(* Tests simple and batch log processors. *)
FUNCTION_BLOCK FB_TestLogProcessors EXTENDS FB_TestSuite

THIS^.testSimpleProcessorExportsEachRecord();
THIS^.testBatchProcessorQueuesAndFlushes();
THIS^.testProcessorsSkipBusyExporter();

(*
	The batch processor queues emitted records in arrival order (oldest at
	the head), dropping the oldest when the queue is full. Flushing moves
	the oldest maxExportBatchSize records into the exporter's queue, on a
	full batch or when the schedule delay elapses, so records leave in order
	and memory stays bounded however fast the PLC logs. queuedCount reports
	the records waiting for export, and droppedCount the records lost.

	FB_LoggerProvider.tick() unstages every processor, so a processor must be
	staged again before each tick.
*)
METHOD testBatchProcessorQueuesAndFlushes : REFERENCE TO FB_Test
VAR
	resourceA: FB_Resource('resource.a');
	resourceB: FB_Resource('resource.b');
	providerA: FB_LoggerProvider(resourceA);
	providerB: FB_LoggerProvider(resourceB);
	scopeA: FB_InstrumentationScope('scope.a', '1.0.0', '');
	scopeB: FB_InstrumentationScope('scope.b', '1.0.0', '');
	loggerAA: FB_Logger(scopeA, providerA);
	loggerAB: FB_Logger(scopeB, providerA);
	loggerBA: FB_Logger(scopeA, providerB);
	exporter: FB_LogRecordExporter_ForInspection;
	processor: FB_LogRecordProcessor_ForBatchInspection(
		maxQueueSize:=10,
		scheduledDelayMillis:=1000,
		maxExportBatchSize:=6,
		exporter:=exporter
	);
	// no exporter, so onEmit only enriches and never queues
	orphanProcessor: FB_LogRecordProcessor_ForBatchInspection(
		maxQueueSize:=10,
		scheduledDelayMillis:=1000,
		maxExportBatchSize:=6,
		exporter:=0
	);
	boundedExporter: FB_LogRecordExporter_ForInspection;
	boundedProcessor: FB_LogRecordProcessor_ForBatchInspection(
		maxQueueSize:=2,
		scheduledDelayMillis:=1000,
		maxExportBatchSize:=3,
		exporter:=boundedExporter
	);
	timerExporter: FB_LogRecordExporter_ForInspection;
	timerProcessor: FB_LogRecordProcessor_ForBatchInspection(
		maxQueueSize:=0,
		scheduledDelayMillis:=0,
		maxExportBatchSize:=3,
		exporter:=timerExporter
	);
	ts1: ULINT := 1;
	ts2: ULINT := 2;
	ts3: ULINT := 3;
	ts4: ULINT := 4;
	ts5: ULINT := 5;
	ts6: ULINT := 6;
	ts7: ULINT := 7;
	ts8: ULINT := 8;
	ts9: ULINT := 9;
	ts10: ULINT := 10;
	ts11: ULINT := 11;
	ts12: ULINT := 12;
	pRec: POINTER TO FB_LogRecord;
END_VAR
TcUnit.TEST('testBatchProcessorQueuesAndFlushes');
	// processor uses maxExportBatchSize 6 so the count-based flush trigger fires without waiting on the timer

	// --- Scenario: records queue in arrival order ---
	// emit interleaved across (resource, scope) pairs
	loggerBA.startLogRecord(severityNumber:=E_SeverityNumber.INFO).setTimestamp(ts1).emit();
	loggerAB.startLogRecord(severityNumber:=E_SeverityNumber.INFO).setTimestamp(ts2).emit();
	loggerAA.startLogRecord(severityNumber:=E_SeverityNumber.INFO).setTimestamp(ts3).emit();
	loggerBA.startLogRecord(severityNumber:=E_SeverityNumber.INFO).setTimestamp(ts4).emit();
	loggerAA.startLogRecord(severityNumber:=E_SeverityNumber.INFO).setTimestamp(ts5).emit();
	// note, it's bad practice to associate processors with multiple providers
	providerA
		.stageProcessor(processor)
		.tick();
	providerB
		.stageProcessor(processor)
		.tick();
	THIS^.AssertTrue(processor.lastOperationSucceeded, 'Expected the last emit to succeed');
	THIS^.AssertEquals_UDINT(5, processor.records.count, 'Expected five queued records');
	THIS^.AssertEquals_UDINT(5, processor.queuedCount, 'Expected queuedCount to report the five queued records');
	THIS^.AssertEquals_UDINT(0, processor.droppedCount, 'Expected droppedCount to be zero before the queue fills');

	// the queue keeps arrival order per provider, oldest at the head
	processor.records.reset();
	pRec := processor.records.next();
	THIS^.AssertTrue(pRec <> 0 AND_THEN pRec^.timestamp = 2, 'Expected queued record 1 to be ts2');
	pRec := processor.records.next();
	THIS^.AssertTrue(pRec <> 0 AND_THEN pRec^.timestamp = 3, 'Expected queued record 2 to be ts3');
	pRec := processor.records.next();
	THIS^.AssertTrue(pRec <> 0 AND_THEN pRec^.timestamp = 5, 'Expected queued record 3 to be ts5');
	pRec := processor.records.next();
	THIS^.AssertTrue(pRec <> 0 AND_THEN pRec^.timestamp = 1, 'Expected queued record 4 to be ts1');
	pRec := processor.records.next();
	THIS^.AssertTrue(pRec <> 0 AND_THEN pRec^.timestamp = 4, 'Expected queued record 5 to be ts4');
	THIS^.AssertTrue(processor.records.next() = 0, 'Expected queue iteration to be exhausted');

	// --- Scenario: a full batch flushes to the exporter in order ---
	// emit one more to reach maxExportBatchSize, triggering a flush
	loggerAB.startLogRecord(severityNumber:=E_SeverityNumber.INFO).setTimestamp(ts6).emit();
	providerA
		.stageProcessor(processor)
		.tick();
	THIS^.AssertEquals_UDINT(0, processor.records.count, 'Expected zero records left after a full batch flush');
	THIS^.AssertEquals_UDINT(0, processor.queuedCount, 'Expected queuedCount to drop to zero once the batch leaves');
	THIS^.AssertEquals_UDINT(6, exporter.records.count, 'Expected six records in the exported batch');

	// exported batch preserves arrival order
	exporter.records.reset();
	pRec := exporter.records.next();
	THIS^.AssertTrue(pRec <> 0 AND_THEN pRec^.timestamp = 2, 'Expected batch record 0 to be ts2');
	pRec := exporter.records.next();
	THIS^.AssertTrue(pRec <> 0 AND_THEN pRec^.timestamp = 3, 'Expected batch record 1 to be ts3');
	pRec := exporter.records.next();
	THIS^.AssertTrue(pRec <> 0 AND_THEN pRec^.timestamp = 5, 'Expected batch record 2 to be ts5');
	pRec := exporter.records.next();
	THIS^.AssertTrue(pRec <> 0 AND_THEN pRec^.timestamp = 1, 'Expected batch record 3 to be ts1');
	pRec := exporter.records.next();
	THIS^.AssertTrue(pRec <> 0 AND_THEN pRec^.timestamp = 4, 'Expected batch record 4 to be ts4');
	pRec := exporter.records.next();
	THIS^.AssertTrue(pRec <> 0 AND_THEN pRec^.timestamp = 6, 'Expected batch record 5 to be ts6');
	THIS^.AssertTrue(exporter.records.next() = 0, 'Expected batch iteration to be exhausted');

	// --- Scenario: a busy exporter holds records in the queue ---
	// the processor still queues records, but no batch leaves
	exporter.busy := TRUE;
	loggerAB.startLogRecord(severityNumber:=E_SeverityNumber.INFO).setTimestamp(ts7).emit();
	providerA
		.stageProcessor(processor)
		.tick();
	THIS^.AssertEquals_UDINT(1, processor.records.count, 'Expected one queued record while the exporter is busy');
	THIS^.AssertEquals_UDINT(6, exporter.records.count, 'Expected the busy exporter to keep the previous batch');

	// --- Scenario: a partial batch waits for the schedule delay ---
	// once free again, the single queued record stays until scheduledDelayMillis (1000 ms) elapses
	exporter.busy := FALSE;
	providerA
		.stageProcessor(processor)
		.tick();
	THIS^.AssertEquals_UDINT(1, processor.records.count, 'Expected the partial batch to wait for the schedule delay');
	THIS^.AssertEquals_UDINT(6, exporter.records.count, 'Expected no new batch before the schedule delay elapses');

	// --- Scenario: no exporter, no queue ---
	// without a bound exporter onEmit only enriches, so nothing is cloned or queued
	loggerAA.startLogRecord(severityNumber:=E_SeverityNumber.INFO).setTimestamp(ts8).emit();
	providerA
		.stageProcessor(orphanProcessor)
		.tick();
	THIS^.AssertEquals_UDINT(0, orphanProcessor.records.count, 'Expected no queued records without a bound exporter');
	THIS^.AssertTrue(orphanProcessor.lastOperationSucceeded, 'Expected onEmit to succeed without a bound exporter');

	// --- Scenario: a full queue drops the oldest record ---
	// boundedProcessor holds 2 records, so the third emit pushes out the first
	THIS^.AssertEquals_UDINT(2, boundedProcessor.records.maxCount, 'Expected the internal queue to be bounded to maxQueueSize');
	loggerAA.startLogRecord(severityNumber:=E_SeverityNumber.INFO).setTimestamp(ts9).emit();
	loggerAB.startLogRecord(severityNumber:=E_SeverityNumber.INFO).setTimestamp(ts10).emit();
	loggerBA.startLogRecord(severityNumber:=E_SeverityNumber.INFO).setTimestamp(ts11).emit();
	providerA
		.stageProcessor(boundedProcessor)
		.tick();
	providerB
		.stageProcessor(boundedProcessor)
		.tick();
	THIS^.AssertEquals_UDINT(2, boundedProcessor.records.count, 'Expected the queue to stay at maxQueueSize');
	THIS^.AssertEquals_UDINT(1, boundedProcessor.records.droppedCount, 'Expected the oldest record to be dropped');
	THIS^.AssertEquals_UDINT(2, boundedProcessor.queuedCount, 'Expected queuedCount to stay at maxQueueSize');
	THIS^.AssertEquals_UDINT(1, boundedProcessor.droppedCount, 'Expected droppedCount to include the evicted record');
	boundedProcessor.records.reset();
	pRec := boundedProcessor.records.next();
	THIS^.AssertTrue(pRec <> 0 AND_THEN pRec^.timestamp = 10, 'Expected ts9 to be dropped and ts10 at the head');
	pRec := boundedProcessor.records.next();
	THIS^.AssertTrue(pRec <> 0 AND_THEN pRec^.timestamp = 11, 'Expected ts11 at the tail');

	// --- Scenario: the schedule timer flushes a partial batch ---
	// timerProcessor has an unbounded queue (maxQueueSize 0) and a 0 ms delay, so one record is enough to flush
	loggerAA.startLogRecord(severityNumber:=E_SeverityNumber.INFO).setTimestamp(ts12).emit();
	providerA
		.stageProcessor(timerProcessor)
		.tick();
	THIS^.AssertEquals_UDINT(0, timerProcessor.records.count, 'Expected the elapsed timer to flush a partial batch');
	THIS^.AssertEquals_UDINT(0, timerProcessor.queuedCount, 'Expected queuedCount to be zero after the timer flush');
	THIS^.AssertEquals_UDINT(1, timerExporter.records.count, 'Expected one record in the timer-triggered batch');
	timerExporter.records.reset();
	pRec := timerExporter.records.next();
	THIS^.AssertTrue(pRec <> 0 AND_THEN pRec^.timestamp = 12, 'Expected the timer-triggered batch record');

	// --- Cleanup: free releases each processor queue ---
	processor.free();
	orphanProcessor.free();
	boundedProcessor.free();
	timerProcessor.free();
	THIS^.AssertTrue(processor.records.count = 0, 'Expected zero records after free');
	THIS^.AssertTrue(orphanProcessor.records.count = 0, 'Expected zero orphan records after free');
	THIS^.AssertTrue(boundedProcessor.records.count = 0, 'Expected zero bounded records after free');
	THIS^.AssertTrue(timerProcessor.records.count = 0, 'Expected zero timer records after free');
TcUnit.TEST_FINISHED();
END_METHOD

(*
	The simple processor hands each emitted record to an idle exporter straight away, as a clone that
	keeps the body, severity and resource snapshot, so the exporter owns a record that outlives the logger's.
*)
METHOD testSimpleProcessorExportsEachRecord : REFERENCE TO FB_Test
VAR
	resource: FB_Resource('');
	provider: FB_LoggerProvider(resource);
	scope: FB_InstrumentationScope('name', 'version', 'schemaUrl');
	logger: FB_Logger(scope, provider);
	exporter: FB_LogRecordExporter_ForInspection;
	processor: FB_LogRecordProcessor_Simple(exporter);
	pRec: POINTER TO FB_LogRecord;
	pBody: POINTER TO FB_String;
END_VAR
TcUnit.TEST('testSimpleProcessorExportsEachRecord');
	resource.attributes.setStringAttribute('plc.name', 'sim.plc');
	logger.startLogRecord(
			severityNumber:=E_SeverityNumber.ERROR
		)
		.setBody('this is a test')
		.emit();
	provider
		.stageProcessor(processor)
		.tick();

	THIS^.AssertEquals_UDINT(1, exporter.records.count, 'Expected the simple processor to export the emitted record');
	exporter.records.reset();
	pRec := exporter.records.next();
	THIS^.AssertTrue(pRec <> 0, 'Expected the exporter to hold the exported record');
	IF pRec <> 0 THEN
		THIS^.AssertTrue(
			pRec^.severityNumber = E_SeverityNumber.ERROR,
			'Expected the exported record to keep its ERROR severity'
		);
		THIS^.AssertTrue(
			pRec^.body <> 0 AND_THEN pRec^.body^.eType = E_ValueType.E_String,
			'Expected the exported record to keep its string body'
		);
		IF pRec^.body <> 0 AND_THEN pRec^.body^.eType = E_ValueType.E_String THEN
			pBody := pRec^.body;
			THIS^.AssertEquals_STRING('this is a test', pBody^.pString^, 'Expected the exported body text');
		END_IF
		THIS^.AssertEquals_UDINT(1, pRec^.resource.attributes.count, 'Expected the exported record to keep the resource attribute');
	END_IF
	exporter.free();
TcUnit.TEST_FINISHED();
END_METHOD

(* Neither processor calls export on a busy exporter, even when the batch processor has a full batch ready. *)
METHOD testProcessorsSkipBusyExporter : REFERENCE TO FB_Test
VAR
	resource: FB_Resource('');
	provider: FB_LoggerProvider(resource);
	scope: FB_InstrumentationScope('scope', '1.0.0', '');
	logger: FB_Logger(scope, provider);
	simpleExporter: FB_LogRecordExporter_ForInspection;
	simpleProcessor: FB_LogRecordProcessor_Simple(simpleExporter);
	batchExporter: FB_LogRecordExporter_ForInspection;
	batchProcessor: FB_LogRecordProcessor_ForBatchInspection(
		maxQueueSize:=10,
		scheduledDelayMillis:=60000,
		maxExportBatchSize:=1,
		exporter:=batchExporter
	);
END_VAR
TcUnit.TEST('testProcessorsSkipBusyExporter');
	simpleExporter.busy := TRUE;
	batchExporter.busy := TRUE;
	logger.startLogRecord(severityNumber:=E_SeverityNumber.INFO).setBody('work').emit();
	provider
		.stageProcessor(simpleProcessor)
		.stageProcessor(batchProcessor)
		.tick();
	THIS^.AssertEquals_UDINT(0, simpleExporter.callsWhileBusy, 'Expected the simple processor not to call a busy exporter');
	THIS^.AssertEquals_UDINT(0, simpleExporter.records.count, 'Expected the busy simple exporter to receive nothing');
	THIS^.AssertEquals_UDINT(0, batchExporter.callsWhileBusy, 'Expected the batch processor not to call a busy exporter');
	THIS^.AssertEquals_UDINT(1, batchProcessor.records.count, 'Expected the full batch to wait in the processor');
	THIS^.AssertEquals_UDINT(1, batchProcessor.queuedCount, 'Expected queuedCount to include the batch held for a busy exporter');
	THIS^.AssertEquals_UDINT(0, batchProcessor.droppedCount, 'Expected a busy exporter not to make the batch processor drop records');

	batchExporter.busy := FALSE;
	provider
		.stageProcessor(batchProcessor)
		.tick();
	THIS^.AssertEquals_UDINT(1, batchExporter.records.count, 'Expected the batch once the exporter is idle');
	THIS^.AssertEquals_UDINT(0, batchProcessor.records.count, 'Expected the processor queue to be empty');
	THIS^.AssertEquals_UDINT(0, batchProcessor.queuedCount, 'Expected queuedCount to be zero once the held batch is exported');
	simpleExporter.free();
	batchExporter.free();
	batchProcessor.free();
TcUnit.TEST_FINISHED();
END_METHOD

END_FUNCTION_BLOCK

(* stored: Version 1.1.0.1
   POU FB_TestLogProcessors: Id {f0aa1fdf-1271-4935-af15-b23605e1dedc}, SpecialFunc None
   Method testBatchProcessorQueuesAndFlushes: Id {7cba4cd6-baeb-4652-979f-3089242ac7bc}
   Method testSimpleProcessorExportsEachRecord: Id {4aa68aa9-8a85-4975-8601-420ccbbed827}
   Method testProcessorsSkipBusyExporter: Id {08a4b76b-58e1-4e23-b2d2-d15472534b6d} *)
